(* IEC 61131-3 sources: STAR-PLC-Agent/results/raw/four_group_20261114/star_deepseek_v2/PUB008/functional/attempt_0001, 1 file *)

(* ---- test_program.st ---- *)
PROGRAM PLC_PRG
VAR
 BenchStep : UDINT := 0;
 BenchCalls : UDINT := 0;
 BenchDone : BOOL := FALSE;
 BenchUut0 : FB_Task;
 BenchUut1 : FB_Task;
 BenchUut2 : FB_Task;
 BenchUut3 : FB_Task;
 BenchUut4 : FB_Task;
 BenchUut5 : FB_Task;
 BenchUut6 : FB_Task;
 BenchUut7 : FB_Task;
 BenchUut8 : FB_Task;
 Binding_0_analogValues : ARRAY[-2..4] OF INT;
 Binding_0_channels : ARRAY[7..13] OF ST_AnalogChannel;
 Binding_1_analogValues : ARRAY[1..5] OF INT;
 Binding_1_channels : ARRAY[1..5] OF ST_AnalogChannel;
 Binding_2_analogValues : ARRAY[1..1] OF INT;
 Binding_2_channels : ARRAY[1..1] OF ST_AnalogChannel;
 Binding_3_analogValues : ARRAY[-3..-3] OF INT;
 Binding_3_channels : ARRAY[9..10] OF ST_AnalogChannel;
 Binding_4_analogValues : ARRAY[-3..-1] OF INT;
 Binding_4_channels : ARRAY[7..9] OF ST_AnalogChannel;
 Binding_5_analogValues : ARRAY[-3..0] OF INT;
 Binding_5_channels : ARRAY[8..9] OF ST_AnalogChannel;
 Binding_6_analogValues : ARRAY[-3..-2] OF INT;
 Binding_6_channels : ARRAY[8..11] OF ST_AnalogChannel;
 Binding_7_analogValues : ARRAY[1..5] OF INT;
 Binding_7_channels : ARRAY[1..5] OF ST_AnalogChannel;
 Binding_8_analogValues : ARRAY[1..5] OF INT;
 Binding_8_channels : ARRAY[1..6] OF ST_AnalogChannel;
 TraceIn_count : ARRAY[0..11] OF DINT;
 TraceOut_analogValues_1 : ARRAY[0..11] OF INT;
 TraceOut_analogValues_2 : ARRAY[0..11] OF INT;
 TraceOut_analogValues_3 : ARRAY[0..11] OF INT;
 TraceOut_analogValues_4 : ARRAY[0..11] OF INT;
 TraceOut_analogValues_5 : ARRAY[0..11] OF INT;
 TraceOut_analogValues_6 : ARRAY[0..11] OF INT;
 TraceOut_analogValues_7 : ARRAY[0..11] OF INT;
 TraceOut_channels_1_enable : ARRAY[0..11] OF BOOL;
 TraceOut_channels_1_hiLIM : ARRAY[0..11] OF REAL;
 TraceOut_channels_1_loLIM : ARRAY[0..11] OF REAL;
 TraceOut_channels_1_bipolar : ARRAY[0..11] OF BOOL;
 TraceOut_channels_1_measuringMode : ARRAY[0..11] OF INT;
 TraceOut_channels_1_retVal : ARRAY[0..11] OF WORD;
 TraceOut_channels_1_outputValue : ARRAY[0..11] OF REAL;
 TraceOut_channels_2_enable : ARRAY[0..11] OF BOOL;
 TraceOut_channels_2_hiLIM : ARRAY[0..11] OF REAL;
 TraceOut_channels_2_loLIM : ARRAY[0..11] OF REAL;
 TraceOut_channels_2_bipolar : ARRAY[0..11] OF BOOL;
 TraceOut_channels_2_measuringMode : ARRAY[0..11] OF INT;
 TraceOut_channels_2_retVal : ARRAY[0..11] OF WORD;
 TraceOut_channels_2_outputValue : ARRAY[0..11] OF REAL;
 TraceOut_channels_3_enable : ARRAY[0..11] OF BOOL;
 TraceOut_channels_3_hiLIM : ARRAY[0..11] OF REAL;
 TraceOut_channels_3_loLIM : ARRAY[0..11] OF REAL;
 TraceOut_channels_3_bipolar : ARRAY[0..11] OF BOOL;
 TraceOut_channels_3_measuringMode : ARRAY[0..11] OF INT;
 TraceOut_channels_3_retVal : ARRAY[0..11] OF WORD;
 TraceOut_channels_3_outputValue : ARRAY[0..11] OF REAL;
 TraceOut_channels_4_enable : ARRAY[0..11] OF BOOL;
 TraceOut_channels_4_hiLIM : ARRAY[0..11] OF REAL;
 TraceOut_channels_4_loLIM : ARRAY[0..11] OF REAL;
 TraceOut_channels_4_bipolar : ARRAY[0..11] OF BOOL;
 TraceOut_channels_4_measuringMode : ARRAY[0..11] OF INT;
 TraceOut_channels_4_retVal : ARRAY[0..11] OF WORD;
 TraceOut_channels_4_outputValue : ARRAY[0..11] OF REAL;
 TraceOut_channels_5_enable : ARRAY[0..11] OF BOOL;
 TraceOut_channels_5_hiLIM : ARRAY[0..11] OF REAL;
 TraceOut_channels_5_loLIM : ARRAY[0..11] OF REAL;
 TraceOut_channels_5_bipolar : ARRAY[0..11] OF BOOL;
 TraceOut_channels_5_measuringMode : ARRAY[0..11] OF INT;
 TraceOut_channels_5_retVal : ARRAY[0..11] OF WORD;
 TraceOut_channels_5_outputValue : ARRAY[0..11] OF REAL;
 TraceOut_channels_6_enable : ARRAY[0..11] OF BOOL;
 TraceOut_channels_6_hiLIM : ARRAY[0..11] OF REAL;
 TraceOut_channels_6_loLIM : ARRAY[0..11] OF REAL;
 TraceOut_channels_6_bipolar : ARRAY[0..11] OF BOOL;
 TraceOut_channels_6_measuringMode : ARRAY[0..11] OF INT;
 TraceOut_channels_6_retVal : ARRAY[0..11] OF WORD;
 TraceOut_channels_6_outputValue : ARRAY[0..11] OF REAL;
 TraceOut_channels_7_enable : ARRAY[0..11] OF BOOL;
 TraceOut_channels_7_hiLIM : ARRAY[0..11] OF REAL;
 TraceOut_channels_7_loLIM : ARRAY[0..11] OF REAL;
 TraceOut_channels_7_bipolar : ARRAY[0..11] OF BOOL;
 TraceOut_channels_7_measuringMode : ARRAY[0..11] OF INT;
 TraceOut_channels_7_retVal : ARRAY[0..11] OF WORD;
 TraceOut_channels_7_outputValue : ARRAY[0..11] OF REAL;
END_VAR

IF NOT BenchDone THEN
 CASE BenchStep OF
 0:
   Binding_0_analogValues[-2] := INT#0;
   Binding_0_analogValues[-1] := INT#27648;
   Binding_0_analogValues[0] := INT#-27648;
   Binding_0_analogValues[1] := INT#0;
   Binding_0_analogValues[2] := INT#27648;
   Binding_0_analogValues[3] := INT#1234;
   Binding_0_analogValues[4] := INT#-1234;
   Binding_0_channels[7].enable := TRUE;
   Binding_0_channels[7].hiLIM := REAL#100.0;
   Binding_0_channels[7].loLIM := REAL#0.0;
   Binding_0_channels[7].bipolar := FALSE;
   Binding_0_channels[7].measuringMode := INT#0;
   Binding_0_channels[7].retVal := WORD#7;
   Binding_0_channels[7].outputValue := REAL#-999.0;
   Binding_0_channels[8].enable := TRUE;
   Binding_0_channels[8].hiLIM := REAL#100.0;
   Binding_0_channels[8].loLIM := REAL#0.0;
   Binding_0_channels[8].bipolar := FALSE;
   Binding_0_channels[8].measuringMode := INT#0;
   Binding_0_channels[8].retVal := WORD#7;
   Binding_0_channels[8].outputValue := REAL#-999.0;
   Binding_0_channels[9].enable := TRUE;
   Binding_0_channels[9].hiLIM := REAL#100.0;
   Binding_0_channels[9].loLIM := REAL#0.0;
   Binding_0_channels[9].bipolar := TRUE;
   Binding_0_channels[9].measuringMode := INT#0;
   Binding_0_channels[9].retVal := WORD#7;
   Binding_0_channels[9].outputValue := REAL#-999.0;
   Binding_0_channels[10].enable := TRUE;
   Binding_0_channels[10].hiLIM := REAL#100.0;
   Binding_0_channels[10].loLIM := REAL#0.0;
   Binding_0_channels[10].bipolar := TRUE;
   Binding_0_channels[10].measuringMode := INT#0;
   Binding_0_channels[10].retVal := WORD#7;
   Binding_0_channels[10].outputValue := REAL#-999.0;
   Binding_0_channels[11].enable := TRUE;
   Binding_0_channels[11].hiLIM := REAL#100.0;
   Binding_0_channels[11].loLIM := REAL#0.0;
   Binding_0_channels[11].bipolar := TRUE;
   Binding_0_channels[11].measuringMode := INT#0;
   Binding_0_channels[11].retVal := WORD#7;
   Binding_0_channels[11].outputValue := REAL#-999.0;
   Binding_0_channels[12].enable := TRUE;
   Binding_0_channels[12].hiLIM := REAL#100.0;
   Binding_0_channels[12].loLIM := REAL#0.0;
   Binding_0_channels[12].bipolar := FALSE;
   Binding_0_channels[12].measuringMode := INT#1;
   Binding_0_channels[12].retVal := WORD#7;
   Binding_0_channels[12].outputValue := REAL#-999.0;
   Binding_0_channels[13].enable := TRUE;
   Binding_0_channels[13].hiLIM := REAL#100.0;
   Binding_0_channels[13].loLIM := REAL#0.0;
   Binding_0_channels[13].bipolar := FALSE;
   Binding_0_channels[13].measuringMode := INT#2;
   Binding_0_channels[13].retVal := WORD#7;
   Binding_0_channels[13].outputValue := REAL#-999.0;
   BenchUut0.count := DINT#7;
   TraceIn_count[0] := BenchUut0.count;
   BenchUut0(analogValues := Binding_0_analogValues, channels := Binding_0_channels);
   TraceOut_analogValues_1[0] := Binding_0_analogValues[-2];
   TraceOut_analogValues_2[0] := Binding_0_analogValues[-1];
   TraceOut_analogValues_3[0] := Binding_0_analogValues[0];
   TraceOut_analogValues_4[0] := Binding_0_analogValues[1];
   TraceOut_analogValues_5[0] := Binding_0_analogValues[2];
   TraceOut_analogValues_6[0] := Binding_0_analogValues[3];
   TraceOut_analogValues_7[0] := Binding_0_analogValues[4];
   TraceOut_channels_1_enable[0] := Binding_0_channels[7].enable;
   TraceOut_channels_1_hiLIM[0] := Binding_0_channels[7].hiLIM;
   TraceOut_channels_1_loLIM[0] := Binding_0_channels[7].loLIM;
   TraceOut_channels_1_bipolar[0] := Binding_0_channels[7].bipolar;
   TraceOut_channels_1_measuringMode[0] := Binding_0_channels[7].measuringMode;
   TraceOut_channels_1_retVal[0] := Binding_0_channels[7].retVal;
   TraceOut_channels_1_outputValue[0] := Binding_0_channels[7].outputValue;
   TraceOut_channels_2_enable[0] := Binding_0_channels[8].enable;
   TraceOut_channels_2_hiLIM[0] := Binding_0_channels[8].hiLIM;
   TraceOut_channels_2_loLIM[0] := Binding_0_channels[8].loLIM;
   TraceOut_channels_2_bipolar[0] := Binding_0_channels[8].bipolar;
   TraceOut_channels_2_measuringMode[0] := Binding_0_channels[8].measuringMode;
   TraceOut_channels_2_retVal[0] := Binding_0_channels[8].retVal;
   TraceOut_channels_2_outputValue[0] := Binding_0_channels[8].outputValue;
   TraceOut_channels_3_enable[0] := Binding_0_channels[9].enable;
   TraceOut_channels_3_hiLIM[0] := Binding_0_channels[9].hiLIM;
   TraceOut_channels_3_loLIM[0] := Binding_0_channels[9].loLIM;
   TraceOut_channels_3_bipolar[0] := Binding_0_channels[9].bipolar;
   TraceOut_channels_3_measuringMode[0] := Binding_0_channels[9].measuringMode;
   TraceOut_channels_3_retVal[0] := Binding_0_channels[9].retVal;
   TraceOut_channels_3_outputValue[0] := Binding_0_channels[9].outputValue;
   TraceOut_channels_4_enable[0] := Binding_0_channels[10].enable;
   TraceOut_channels_4_hiLIM[0] := Binding_0_channels[10].hiLIM;
   TraceOut_channels_4_loLIM[0] := Binding_0_channels[10].loLIM;
   TraceOut_channels_4_bipolar[0] := Binding_0_channels[10].bipolar;
   TraceOut_channels_4_measuringMode[0] := Binding_0_channels[10].measuringMode;
   TraceOut_channels_4_retVal[0] := Binding_0_channels[10].retVal;
   TraceOut_channels_4_outputValue[0] := Binding_0_channels[10].outputValue;
   TraceOut_channels_5_enable[0] := Binding_0_channels[11].enable;
   TraceOut_channels_5_hiLIM[0] := Binding_0_channels[11].hiLIM;
   TraceOut_channels_5_loLIM[0] := Binding_0_channels[11].loLIM;
   TraceOut_channels_5_bipolar[0] := Binding_0_channels[11].bipolar;
   TraceOut_channels_5_measuringMode[0] := Binding_0_channels[11].measuringMode;
   TraceOut_channels_5_retVal[0] := Binding_0_channels[11].retVal;
   TraceOut_channels_5_outputValue[0] := Binding_0_channels[11].outputValue;
   TraceOut_channels_6_enable[0] := Binding_0_channels[12].enable;
   TraceOut_channels_6_hiLIM[0] := Binding_0_channels[12].hiLIM;
   TraceOut_channels_6_loLIM[0] := Binding_0_channels[12].loLIM;
   TraceOut_channels_6_bipolar[0] := Binding_0_channels[12].bipolar;
   TraceOut_channels_6_measuringMode[0] := Binding_0_channels[12].measuringMode;
   TraceOut_channels_6_retVal[0] := Binding_0_channels[12].retVal;
   TraceOut_channels_6_outputValue[0] := Binding_0_channels[12].outputValue;
   TraceOut_channels_7_enable[0] := Binding_0_channels[13].enable;
   TraceOut_channels_7_hiLIM[0] := Binding_0_channels[13].hiLIM;
   TraceOut_channels_7_loLIM[0] := Binding_0_channels[13].loLIM;
   TraceOut_channels_7_bipolar[0] := Binding_0_channels[13].bipolar;
   TraceOut_channels_7_measuringMode[0] := Binding_0_channels[13].measuringMode;
   TraceOut_channels_7_retVal[0] := Binding_0_channels[13].retVal;
   TraceOut_channels_7_outputValue[0] := Binding_0_channels[13].outputValue;
   BenchCalls := BenchCalls + 1;
 1:
   Binding_1_analogValues[1] := INT#1;
   Binding_1_analogValues[2] := INT#2;
   Binding_1_analogValues[3] := INT#3;
   Binding_1_analogValues[4] := INT#4;
   Binding_1_analogValues[5] := INT#5;
   Binding_1_channels[1].enable := FALSE;
   Binding_1_channels[1].hiLIM := REAL#100.0;
   Binding_1_channels[1].loLIM := REAL#0.0;
   Binding_1_channels[1].bipolar := FALSE;
   Binding_1_channels[1].measuringMode := INT#0;
   Binding_1_channels[1].retVal := WORD#7;
   Binding_1_channels[1].outputValue := REAL#-999.0;
   Binding_1_channels[2].enable := TRUE;
   Binding_1_channels[2].hiLIM := REAL#0.0;
   Binding_1_channels[2].loLIM := REAL#10.0;
   Binding_1_channels[2].bipolar := FALSE;
   Binding_1_channels[2].measuringMode := INT#9;
   Binding_1_channels[2].retVal := WORD#7;
   Binding_1_channels[2].outputValue := REAL#-999.0;
   Binding_1_channels[3].enable := TRUE;
   Binding_1_channels[3].hiLIM := REAL#10.0;
   Binding_1_channels[3].loLIM := REAL#10.0;
   Binding_1_channels[3].bipolar := FALSE;
   Binding_1_channels[3].measuringMode := INT#0;
   Binding_1_channels[3].retVal := WORD#7;
   Binding_1_channels[3].outputValue := REAL#-999.0;
   Binding_1_channels[4].enable := TRUE;
   Binding_1_channels[4].hiLIM := REAL#100.0;
   Binding_1_channels[4].loLIM := REAL#0.0;
   Binding_1_channels[4].bipolar := FALSE;
   Binding_1_channels[4].measuringMode := INT#2;
   Binding_1_channels[4].retVal := WORD#7;
   Binding_1_channels[4].outputValue := REAL#-999.0;
   Binding_1_channels[5].enable := TRUE;
   Binding_1_channels[5].hiLIM := REAL#100.0;
   Binding_1_channels[5].loLIM := REAL#0.0;
   Binding_1_channels[5].bipolar := FALSE;
   Binding_1_channels[5].measuringMode := INT#0;
   Binding_1_channels[5].retVal := WORD#7;
   Binding_1_channels[5].outputValue := REAL#-999.0;
   BenchUut1.count := DINT#4;
   TraceIn_count[1] := BenchUut1.count;
   BenchUut1(analogValues := Binding_1_analogValues, channels := Binding_1_channels);
   TraceOut_analogValues_1[1] := Binding_1_analogValues[1];
   TraceOut_analogValues_2[1] := Binding_1_analogValues[2];
   TraceOut_analogValues_3[1] := Binding_1_analogValues[3];
   TraceOut_analogValues_4[1] := Binding_1_analogValues[4];
   TraceOut_analogValues_5[1] := Binding_1_analogValues[5];
   TraceOut_channels_1_enable[1] := Binding_1_channels[1].enable;
   TraceOut_channels_1_hiLIM[1] := Binding_1_channels[1].hiLIM;
   TraceOut_channels_1_loLIM[1] := Binding_1_channels[1].loLIM;
   TraceOut_channels_1_bipolar[1] := Binding_1_channels[1].bipolar;
   TraceOut_channels_1_measuringMode[1] := Binding_1_channels[1].measuringMode;
   TraceOut_channels_1_retVal[1] := Binding_1_channels[1].retVal;
   TraceOut_channels_1_outputValue[1] := Binding_1_channels[1].outputValue;
   TraceOut_channels_2_enable[1] := Binding_1_channels[2].enable;
   TraceOut_channels_2_hiLIM[1] := Binding_1_channels[2].hiLIM;
   TraceOut_channels_2_loLIM[1] := Binding_1_channels[2].loLIM;
   TraceOut_channels_2_bipolar[1] := Binding_1_channels[2].bipolar;
   TraceOut_channels_2_measuringMode[1] := Binding_1_channels[2].measuringMode;
   TraceOut_channels_2_retVal[1] := Binding_1_channels[2].retVal;
   TraceOut_channels_2_outputValue[1] := Binding_1_channels[2].outputValue;
   TraceOut_channels_3_enable[1] := Binding_1_channels[3].enable;
   TraceOut_channels_3_hiLIM[1] := Binding_1_channels[3].hiLIM;
   TraceOut_channels_3_loLIM[1] := Binding_1_channels[3].loLIM;
   TraceOut_channels_3_bipolar[1] := Binding_1_channels[3].bipolar;
   TraceOut_channels_3_measuringMode[1] := Binding_1_channels[3].measuringMode;
   TraceOut_channels_3_retVal[1] := Binding_1_channels[3].retVal;
   TraceOut_channels_3_outputValue[1] := Binding_1_channels[3].outputValue;
   TraceOut_channels_4_enable[1] := Binding_1_channels[4].enable;
   TraceOut_channels_4_hiLIM[1] := Binding_1_channels[4].hiLIM;
   TraceOut_channels_4_loLIM[1] := Binding_1_channels[4].loLIM;
   TraceOut_channels_4_bipolar[1] := Binding_1_channels[4].bipolar;
   TraceOut_channels_4_measuringMode[1] := Binding_1_channels[4].measuringMode;
   TraceOut_channels_4_retVal[1] := Binding_1_channels[4].retVal;
   TraceOut_channels_4_outputValue[1] := Binding_1_channels[4].outputValue;
   TraceOut_channels_5_enable[1] := Binding_1_channels[5].enable;
   TraceOut_channels_5_hiLIM[1] := Binding_1_channels[5].hiLIM;
   TraceOut_channels_5_loLIM[1] := Binding_1_channels[5].loLIM;
   TraceOut_channels_5_bipolar[1] := Binding_1_channels[5].bipolar;
   TraceOut_channels_5_measuringMode[1] := Binding_1_channels[5].measuringMode;
   TraceOut_channels_5_retVal[1] := Binding_1_channels[5].retVal;
   TraceOut_channels_5_outputValue[1] := Binding_1_channels[5].outputValue;
   BenchCalls := BenchCalls + 1;
 2:
   Binding_2_analogValues[1] := INT#-27648;
   Binding_2_channels[1].enable := TRUE;
   Binding_2_channels[1].hiLIM := REAL#100.0;
   Binding_2_channels[1].loLIM := REAL#0.0;
   Binding_2_channels[1].bipolar := FALSE;
   Binding_2_channels[1].measuringMode := INT#0;
   Binding_2_channels[1].retVal := WORD#7;
   Binding_2_channels[1].outputValue := REAL#-999.0;
   BenchUut2.count := DINT#0;
   TraceIn_count[2] := BenchUut2.count;
   BenchUut2(analogValues := Binding_2_analogValues, channels := Binding_2_channels);
   TraceOut_analogValues_1[2] := Binding_2_analogValues[1];
   TraceOut_channels_1_enable[2] := Binding_2_channels[1].enable;
   TraceOut_channels_1_hiLIM[2] := Binding_2_channels[1].hiLIM;
   TraceOut_channels_1_loLIM[2] := Binding_2_channels[1].loLIM;
   TraceOut_channels_1_bipolar[2] := Binding_2_channels[1].bipolar;
   TraceOut_channels_1_measuringMode[2] := Binding_2_channels[1].measuringMode;
   TraceOut_channels_1_retVal[2] := Binding_2_channels[1].retVal;
   TraceOut_channels_1_outputValue[2] := Binding_2_channels[1].outputValue;
   BenchCalls := BenchCalls + 1;
 3:
   Binding_2_analogValues[1] := INT#-27648;
   Binding_2_channels[1].enable := TRUE;
   Binding_2_channels[1].hiLIM := REAL#100.0;
   Binding_2_channels[1].loLIM := REAL#0.0;
   Binding_2_channels[1].bipolar := FALSE;
   Binding_2_channels[1].measuringMode := INT#0;
   Binding_2_channels[1].retVal := WORD#7;
   Binding_2_channels[1].outputValue := REAL#-999.0;
   BenchUut2.count := DINT#1;
   TraceIn_count[3] := BenchUut2.count;
   BenchUut2(analogValues := Binding_2_analogValues, channels := Binding_2_channels);
   TraceOut_analogValues_1[3] := Binding_2_analogValues[1];
   TraceOut_channels_1_enable[3] := Binding_2_channels[1].enable;
   TraceOut_channels_1_hiLIM[3] := Binding_2_channels[1].hiLIM;
   TraceOut_channels_1_loLIM[3] := Binding_2_channels[1].loLIM;
   TraceOut_channels_1_bipolar[3] := Binding_2_channels[1].bipolar;
   TraceOut_channels_1_measuringMode[3] := Binding_2_channels[1].measuringMode;
   TraceOut_channels_1_retVal[3] := Binding_2_channels[1].retVal;
   TraceOut_channels_1_outputValue[3] := Binding_2_channels[1].outputValue;
   BenchCalls := BenchCalls + 1;
 4:
   Binding_3_analogValues[-3] := INT#32767;
   Binding_3_channels[9].enable := TRUE;
   Binding_3_channels[9].hiLIM := REAL#27648.0;
   Binding_3_channels[9].loLIM := REAL#-27648.0;
   Binding_3_channels[9].bipolar := TRUE;
   Binding_3_channels[9].measuringMode := INT#0;
   Binding_3_channels[9].retVal := WORD#7;
   Binding_3_channels[9].outputValue := REAL#-999.0;
   Binding_3_channels[10].enable := TRUE;
   Binding_3_channels[10].hiLIM := REAL#27648.0;
   Binding_3_channels[10].loLIM := REAL#-27648.0;
   Binding_3_channels[10].bipolar := TRUE;
   Binding_3_channels[10].measuringMode := INT#0;
   Binding_3_channels[10].retVal := WORD#7;
   Binding_3_channels[10].outputValue := REAL#33.0;
   BenchUut3.count := DINT#1;
   TraceIn_count[4] := BenchUut3.count;
   BenchUut3(analogValues := Binding_3_analogValues, channels := Binding_3_channels);
   TraceOut_analogValues_1[4] := Binding_3_analogValues[-3];
   TraceOut_channels_1_enable[4] := Binding_3_channels[9].enable;
   TraceOut_channels_1_hiLIM[4] := Binding_3_channels[9].hiLIM;
   TraceOut_channels_1_loLIM[4] := Binding_3_channels[9].loLIM;
   TraceOut_channels_1_bipolar[4] := Binding_3_channels[9].bipolar;
   TraceOut_channels_1_measuringMode[4] := Binding_3_channels[9].measuringMode;
   TraceOut_channels_1_retVal[4] := Binding_3_channels[9].retVal;
   TraceOut_channels_1_outputValue[4] := Binding_3_channels[9].outputValue;
   TraceOut_channels_2_enable[4] := Binding_3_channels[10].enable;
   TraceOut_channels_2_hiLIM[4] := Binding_3_channels[10].hiLIM;
   TraceOut_channels_2_loLIM[4] := Binding_3_channels[10].loLIM;
   TraceOut_channels_2_bipolar[4] := Binding_3_channels[10].bipolar;
   TraceOut_channels_2_measuringMode[4] := Binding_3_channels[10].measuringMode;
   TraceOut_channels_2_retVal[4] := Binding_3_channels[10].retVal;
   TraceOut_channels_2_outputValue[4] := Binding_3_channels[10].outputValue;
   BenchCalls := BenchCalls + 1;
 5:
   Binding_4_analogValues[-3] := INT#1000;
   Binding_4_analogValues[-2] := INT#-1000;
   Binding_4_analogValues[-1] := INT#30000;
   Binding_4_channels[7].enable := FALSE;
   Binding_4_channels[7].hiLIM := REAL#0.0;
   Binding_4_channels[7].loLIM := REAL#100.0;
   Binding_4_channels[7].bipolar := FALSE;
   Binding_4_channels[7].measuringMode := INT#9;
   Binding_4_channels[7].retVal := WORD#123;
   Binding_4_channels[7].outputValue := REAL#-42.5;
   Binding_4_channels[8].enable := TRUE;
   Binding_4_channels[8].hiLIM := REAL#5.0;
   Binding_4_channels[8].loLIM := REAL#5.0;
   Binding_4_channels[8].bipolar := FALSE;
   Binding_4_channels[8].measuringMode := INT#1;
   Binding_4_channels[8].retVal := WORD#0;
   Binding_4_channels[8].outputValue := REAL#12.25;
   Binding_4_channels[9].enable := TRUE;
   Binding_4_channels[9].hiLIM := REAL#100.0;
   Binding_4_channels[9].loLIM := REAL#0.0;
   Binding_4_channels[9].bipolar := FALSE;
   Binding_4_channels[9].measuringMode := INT#0;
   Binding_4_channels[9].retVal := WORD#0;
   Binding_4_channels[9].outputValue := REAL#0.0;
   BenchUut4.count := DINT#3;
   TraceIn_count[5] := BenchUut4.count;
   BenchUut4(analogValues := Binding_4_analogValues, channels := Binding_4_channels);
   TraceOut_analogValues_1[5] := Binding_4_analogValues[-3];
   TraceOut_analogValues_2[5] := Binding_4_analogValues[-2];
   TraceOut_analogValues_3[5] := Binding_4_analogValues[-1];
   TraceOut_channels_1_enable[5] := Binding_4_channels[7].enable;
   TraceOut_channels_1_hiLIM[5] := Binding_4_channels[7].hiLIM;
   TraceOut_channels_1_loLIM[5] := Binding_4_channels[7].loLIM;
   TraceOut_channels_1_bipolar[5] := Binding_4_channels[7].bipolar;
   TraceOut_channels_1_measuringMode[5] := Binding_4_channels[7].measuringMode;
   TraceOut_channels_1_retVal[5] := Binding_4_channels[7].retVal;
   TraceOut_channels_1_outputValue[5] := Binding_4_channels[7].outputValue;
   TraceOut_channels_2_enable[5] := Binding_4_channels[8].enable;
   TraceOut_channels_2_hiLIM[5] := Binding_4_channels[8].hiLIM;
   TraceOut_channels_2_loLIM[5] := Binding_4_channels[8].loLIM;
   TraceOut_channels_2_bipolar[5] := Binding_4_channels[8].bipolar;
   TraceOut_channels_2_measuringMode[5] := Binding_4_channels[8].measuringMode;
   TraceOut_channels_2_retVal[5] := Binding_4_channels[8].retVal;
   TraceOut_channels_2_outputValue[5] := Binding_4_channels[8].outputValue;
   TraceOut_channels_3_enable[5] := Binding_4_channels[9].enable;
   TraceOut_channels_3_hiLIM[5] := Binding_4_channels[9].hiLIM;
   TraceOut_channels_3_loLIM[5] := Binding_4_channels[9].loLIM;
   TraceOut_channels_3_bipolar[5] := Binding_4_channels[9].bipolar;
   TraceOut_channels_3_measuringMode[5] := Binding_4_channels[9].measuringMode;
   TraceOut_channels_3_retVal[5] := Binding_4_channels[9].retVal;
   TraceOut_channels_3_outputValue[5] := Binding_4_channels[9].outputValue;
   BenchCalls := BenchCalls + 1;
 6:
   Binding_4_analogValues[-3] := INT#-30000;
   Binding_4_analogValues[-2] := INT#1234;
   Binding_4_analogValues[-1] := INT#0;
   Binding_4_analogValues[0] := INT#999;
   Binding_4_channels[7].enable := TRUE;
   Binding_4_channels[7].hiLIM := REAL#10.0;
   Binding_4_channels[7].loLIM := REAL#-10.0;
   Binding_4_channels[7].bipolar := FALSE;
   Binding_4_channels[7].measuringMode := INT#2;
   Binding_4_channels[7].retVal := WORD#0;
   Binding_4_channels[7].outputValue := REAL#1.0;
   Binding_4_channels[8].enable := TRUE;
   Binding_4_channels[8].hiLIM := REAL#10.0;
   Binding_4_channels[8].loLIM := REAL#20.0;
   Binding_4_channels[8].bipolar := FALSE;
   Binding_4_channels[8].measuringMode := INT#2;
   Binding_4_channels[8].retVal := WORD#0;
   Binding_4_channels[8].outputValue := REAL#3.5;
   Binding_4_channels[9].enable := TRUE;
   Binding_4_channels[9].hiLIM := REAL#10.0;
   Binding_4_channels[9].loLIM := REAL#0.0;
   Binding_4_channels[9].bipolar := TRUE;
   Binding_4_channels[9].measuringMode := INT#0;
   Binding_4_channels[9].retVal := WORD#0;
   Binding_4_channels[9].outputValue := REAL#0.0;
   BenchUut4.count := DINT#3;
   TraceIn_count[6] := BenchUut4.count;
   BenchUut4(analogValues := Binding_4_analogValues, channels := Binding_4_channels);
   TraceOut_analogValues_1[6] := Binding_4_analogValues[-3];
   TraceOut_analogValues_2[6] := Binding_4_analogValues[-2];
   TraceOut_analogValues_3[6] := Binding_4_analogValues[-1];
   TraceOut_analogValues_4[6] := Binding_4_analogValues[0];
   TraceOut_channels_1_enable[6] := Binding_4_channels[7].enable;
   TraceOut_channels_1_hiLIM[6] := Binding_4_channels[7].hiLIM;
   TraceOut_channels_1_loLIM[6] := Binding_4_channels[7].loLIM;
   TraceOut_channels_1_bipolar[6] := Binding_4_channels[7].bipolar;
   TraceOut_channels_1_measuringMode[6] := Binding_4_channels[7].measuringMode;
   TraceOut_channels_1_retVal[6] := Binding_4_channels[7].retVal;
   TraceOut_channels_1_outputValue[6] := Binding_4_channels[7].outputValue;
   TraceOut_channels_2_enable[6] := Binding_4_channels[8].enable;
   TraceOut_channels_2_hiLIM[6] := Binding_4_channels[8].hiLIM;
   TraceOut_channels_2_loLIM[6] := Binding_4_channels[8].loLIM;
   TraceOut_channels_2_bipolar[6] := Binding_4_channels[8].bipolar;
   TraceOut_channels_2_measuringMode[6] := Binding_4_channels[8].measuringMode;
   TraceOut_channels_2_retVal[6] := Binding_4_channels[8].retVal;
   TraceOut_channels_2_outputValue[6] := Binding_4_channels[8].outputValue;
   TraceOut_channels_3_enable[6] := Binding_4_channels[9].enable;
   TraceOut_channels_3_hiLIM[6] := Binding_4_channels[9].hiLIM;
   TraceOut_channels_3_loLIM[6] := Binding_4_channels[9].loLIM;
   TraceOut_channels_3_bipolar[6] := Binding_4_channels[9].bipolar;
   TraceOut_channels_3_measuringMode[6] := Binding_4_channels[9].measuringMode;
   TraceOut_channels_3_retVal[6] := Binding_4_channels[9].retVal;
   TraceOut_channels_3_outputValue[6] := Binding_4_channels[9].outputValue;
   BenchCalls := BenchCalls + 1;
 7:
   Binding_5_analogValues[-3] := INT#0;
   Binding_5_analogValues[-2] := INT#27648;
   Binding_5_analogValues[-1] := INT#-27648;
   Binding_5_analogValues[0] := INT#0;
   Binding_5_channels[8].enable := TRUE;
   Binding_5_channels[8].hiLIM := REAL#100.0;
   Binding_5_channels[8].loLIM := REAL#0.0;
   Binding_5_channels[8].bipolar := FALSE;
   Binding_5_channels[8].measuringMode := INT#0;
   Binding_5_channels[8].retVal := WORD#7;
   Binding_5_channels[8].outputValue := REAL#-999.0;
   Binding_5_channels[9].enable := TRUE;
   Binding_5_channels[9].hiLIM := REAL#100.0;
   Binding_5_channels[9].loLIM := REAL#0.0;
   Binding_5_channels[9].bipolar := FALSE;
   Binding_5_channels[9].measuringMode := INT#0;
   Binding_5_channels[9].retVal := WORD#7;
   Binding_5_channels[9].outputValue := REAL#-999.0;
   BenchUut5.count := DINT#2;
   TraceIn_count[7] := BenchUut5.count;
   BenchUut5(analogValues := Binding_5_analogValues, channels := Binding_5_channels);
   TraceOut_analogValues_1[7] := Binding_5_analogValues[-3];
   TraceOut_analogValues_2[7] := Binding_5_analogValues[-2];
   TraceOut_analogValues_3[7] := Binding_5_analogValues[-1];
   TraceOut_analogValues_4[7] := Binding_5_analogValues[0];
   TraceOut_channels_1_enable[7] := Binding_5_channels[8].enable;
   TraceOut_channels_1_hiLIM[7] := Binding_5_channels[8].hiLIM;
   TraceOut_channels_1_loLIM[7] := Binding_5_channels[8].loLIM;
   TraceOut_channels_1_bipolar[7] := Binding_5_channels[8].bipolar;
   TraceOut_channels_1_measuringMode[7] := Binding_5_channels[8].measuringMode;
   TraceOut_channels_1_retVal[7] := Binding_5_channels[8].retVal;
   TraceOut_channels_1_outputValue[7] := Binding_5_channels[8].outputValue;
   TraceOut_channels_2_enable[7] := Binding_5_channels[9].enable;
   TraceOut_channels_2_hiLIM[7] := Binding_5_channels[9].hiLIM;
   TraceOut_channels_2_loLIM[7] := Binding_5_channels[9].loLIM;
   TraceOut_channels_2_bipolar[7] := Binding_5_channels[9].bipolar;
   TraceOut_channels_2_measuringMode[7] := Binding_5_channels[9].measuringMode;
   TraceOut_channels_2_retVal[7] := Binding_5_channels[9].retVal;
   TraceOut_channels_2_outputValue[7] := Binding_5_channels[9].outputValue;
   BenchCalls := BenchCalls + 1;
 8:
   Binding_6_analogValues[-3] := INT#0;
   Binding_6_analogValues[-2] := INT#27648;
   Binding_6_channels[8].enable := TRUE;
   Binding_6_channels[8].hiLIM := REAL#100.0;
   Binding_6_channels[8].loLIM := REAL#0.0;
   Binding_6_channels[8].bipolar := FALSE;
   Binding_6_channels[8].measuringMode := INT#0;
   Binding_6_channels[8].retVal := WORD#7;
   Binding_6_channels[8].outputValue := REAL#-999.0;
   Binding_6_channels[9].enable := TRUE;
   Binding_6_channels[9].hiLIM := REAL#100.0;
   Binding_6_channels[9].loLIM := REAL#0.0;
   Binding_6_channels[9].bipolar := FALSE;
   Binding_6_channels[9].measuringMode := INT#0;
   Binding_6_channels[9].retVal := WORD#7;
   Binding_6_channels[9].outputValue := REAL#-999.0;
   Binding_6_channels[10].enable := TRUE;
   Binding_6_channels[10].hiLIM := REAL#100.0;
   Binding_6_channels[10].loLIM := REAL#0.0;
   Binding_6_channels[10].bipolar := TRUE;
   Binding_6_channels[10].measuringMode := INT#0;
   Binding_6_channels[10].retVal := WORD#7;
   Binding_6_channels[10].outputValue := REAL#-999.0;
   Binding_6_channels[11].enable := TRUE;
   Binding_6_channels[11].hiLIM := REAL#100.0;
   Binding_6_channels[11].loLIM := REAL#0.0;
   Binding_6_channels[11].bipolar := TRUE;
   Binding_6_channels[11].measuringMode := INT#0;
   Binding_6_channels[11].retVal := WORD#7;
   Binding_6_channels[11].outputValue := REAL#-999.0;
   BenchUut6.count := DINT#2;
   TraceIn_count[8] := BenchUut6.count;
   BenchUut6(analogValues := Binding_6_analogValues, channels := Binding_6_channels);
   TraceOut_analogValues_1[8] := Binding_6_analogValues[-3];
   TraceOut_analogValues_2[8] := Binding_6_analogValues[-2];
   TraceOut_channels_1_enable[8] := Binding_6_channels[8].enable;
   TraceOut_channels_1_hiLIM[8] := Binding_6_channels[8].hiLIM;
   TraceOut_channels_1_loLIM[8] := Binding_6_channels[8].loLIM;
   TraceOut_channels_1_bipolar[8] := Binding_6_channels[8].bipolar;
   TraceOut_channels_1_measuringMode[8] := Binding_6_channels[8].measuringMode;
   TraceOut_channels_1_retVal[8] := Binding_6_channels[8].retVal;
   TraceOut_channels_1_outputValue[8] := Binding_6_channels[8].outputValue;
   TraceOut_channels_2_enable[8] := Binding_6_channels[9].enable;
   TraceOut_channels_2_hiLIM[8] := Binding_6_channels[9].hiLIM;
   TraceOut_channels_2_loLIM[8] := Binding_6_channels[9].loLIM;
   TraceOut_channels_2_bipolar[8] := Binding_6_channels[9].bipolar;
   TraceOut_channels_2_measuringMode[8] := Binding_6_channels[9].measuringMode;
   TraceOut_channels_2_retVal[8] := Binding_6_channels[9].retVal;
   TraceOut_channels_2_outputValue[8] := Binding_6_channels[9].outputValue;
   TraceOut_channels_3_enable[8] := Binding_6_channels[10].enable;
   TraceOut_channels_3_hiLIM[8] := Binding_6_channels[10].hiLIM;
   TraceOut_channels_3_loLIM[8] := Binding_6_channels[10].loLIM;
   TraceOut_channels_3_bipolar[8] := Binding_6_channels[10].bipolar;
   TraceOut_channels_3_measuringMode[8] := Binding_6_channels[10].measuringMode;
   TraceOut_channels_3_retVal[8] := Binding_6_channels[10].retVal;
   TraceOut_channels_3_outputValue[8] := Binding_6_channels[10].outputValue;
   TraceOut_channels_4_enable[8] := Binding_6_channels[11].enable;
   TraceOut_channels_4_hiLIM[8] := Binding_6_channels[11].hiLIM;
   TraceOut_channels_4_loLIM[8] := Binding_6_channels[11].loLIM;
   TraceOut_channels_4_bipolar[8] := Binding_6_channels[11].bipolar;
   TraceOut_channels_4_measuringMode[8] := Binding_6_channels[11].measuringMode;
   TraceOut_channels_4_retVal[8] := Binding_6_channels[11].retVal;
   TraceOut_channels_4_outputValue[8] := Binding_6_channels[11].outputValue;
   BenchCalls := BenchCalls + 1;
 9:
   Binding_7_analogValues[1] := INT#27648;
   Binding_7_analogValues[2] := INT#13824;
   Binding_7_analogValues[3] := INT#27648;
   Binding_7_analogValues[4] := INT#27648;
   Binding_7_analogValues[5] := INT#500;
   Binding_7_channels[1].enable := TRUE;
   Binding_7_channels[1].hiLIM := REAL#100.0;
   Binding_7_channels[1].loLIM := REAL#0.0;
   Binding_7_channels[1].bipolar := FALSE;
   Binding_7_channels[1].measuringMode := INT#0;
   Binding_7_channels[1].retVal := WORD#7;
   Binding_7_channels[1].outputValue := REAL#-999.0;
   Binding_7_channels[2].enable := TRUE;
   Binding_7_channels[2].hiLIM := REAL#50.0;
   Binding_7_channels[2].loLIM := REAL#-50.0;
   Binding_7_channels[2].bipolar := FALSE;
   Binding_7_channels[2].measuringMode := INT#0;
   Binding_7_channels[2].retVal := WORD#7;
   Binding_7_channels[2].outputValue := REAL#-999.0;
   Binding_7_channels[3].enable := TRUE;
   Binding_7_channels[3].hiLIM := REAL#100.0;
   Binding_7_channels[3].loLIM := REAL#0.0;
   Binding_7_channels[3].bipolar := FALSE;
   Binding_7_channels[3].measuringMode := INT#0;
   Binding_7_channels[3].retVal := WORD#7;
   Binding_7_channels[3].outputValue := REAL#-999.0;
   Binding_7_channels[4].enable := TRUE;
   Binding_7_channels[4].hiLIM := REAL#100.0;
   Binding_7_channels[4].loLIM := REAL#0.0;
   Binding_7_channels[4].bipolar := FALSE;
   Binding_7_channels[4].measuringMode := INT#0;
   Binding_7_channels[4].retVal := WORD#7;
   Binding_7_channels[4].outputValue := REAL#-999.0;
   Binding_7_channels[5].enable := TRUE;
   Binding_7_channels[5].hiLIM := REAL#100.0;
   Binding_7_channels[5].loLIM := REAL#0.0;
   Binding_7_channels[5].bipolar := FALSE;
   Binding_7_channels[5].measuringMode := INT#1;
   Binding_7_channels[5].retVal := WORD#7;
   Binding_7_channels[5].outputValue := REAL#-999.0;
   BenchUut7.count := DINT#5;
   TraceIn_count[9] := BenchUut7.count;
   BenchUut7(analogValues := Binding_7_analogValues, channels := Binding_7_channels);
   TraceOut_analogValues_1[9] := Binding_7_analogValues[1];
   TraceOut_analogValues_2[9] := Binding_7_analogValues[2];
   TraceOut_analogValues_3[9] := Binding_7_analogValues[3];
   TraceOut_analogValues_4[9] := Binding_7_analogValues[4];
   TraceOut_analogValues_5[9] := Binding_7_analogValues[5];
   TraceOut_channels_1_enable[9] := Binding_7_channels[1].enable;
   TraceOut_channels_1_hiLIM[9] := Binding_7_channels[1].hiLIM;
   TraceOut_channels_1_loLIM[9] := Binding_7_channels[1].loLIM;
   TraceOut_channels_1_bipolar[9] := Binding_7_channels[1].bipolar;
   TraceOut_channels_1_measuringMode[9] := Binding_7_channels[1].measuringMode;
   TraceOut_channels_1_retVal[9] := Binding_7_channels[1].retVal;
   TraceOut_channels_1_outputValue[9] := Binding_7_channels[1].outputValue;
   TraceOut_channels_2_enable[9] := Binding_7_channels[2].enable;
   TraceOut_channels_2_hiLIM[9] := Binding_7_channels[2].hiLIM;
   TraceOut_channels_2_loLIM[9] := Binding_7_channels[2].loLIM;
   TraceOut_channels_2_bipolar[9] := Binding_7_channels[2].bipolar;
   TraceOut_channels_2_measuringMode[9] := Binding_7_channels[2].measuringMode;
   TraceOut_channels_2_retVal[9] := Binding_7_channels[2].retVal;
   TraceOut_channels_2_outputValue[9] := Binding_7_channels[2].outputValue;
   TraceOut_channels_3_enable[9] := Binding_7_channels[3].enable;
   TraceOut_channels_3_hiLIM[9] := Binding_7_channels[3].hiLIM;
   TraceOut_channels_3_loLIM[9] := Binding_7_channels[3].loLIM;
   TraceOut_channels_3_bipolar[9] := Binding_7_channels[3].bipolar;
   TraceOut_channels_3_measuringMode[9] := Binding_7_channels[3].measuringMode;
   TraceOut_channels_3_retVal[9] := Binding_7_channels[3].retVal;
   TraceOut_channels_3_outputValue[9] := Binding_7_channels[3].outputValue;
   TraceOut_channels_4_enable[9] := Binding_7_channels[4].enable;
   TraceOut_channels_4_hiLIM[9] := Binding_7_channels[4].hiLIM;
   TraceOut_channels_4_loLIM[9] := Binding_7_channels[4].loLIM;
   TraceOut_channels_4_bipolar[9] := Binding_7_channels[4].bipolar;
   TraceOut_channels_4_measuringMode[9] := Binding_7_channels[4].measuringMode;
   TraceOut_channels_4_retVal[9] := Binding_7_channels[4].retVal;
   TraceOut_channels_4_outputValue[9] := Binding_7_channels[4].outputValue;
   TraceOut_channels_5_enable[9] := Binding_7_channels[5].enable;
   TraceOut_channels_5_hiLIM[9] := Binding_7_channels[5].hiLIM;
   TraceOut_channels_5_loLIM[9] := Binding_7_channels[5].loLIM;
   TraceOut_channels_5_bipolar[9] := Binding_7_channels[5].bipolar;
   TraceOut_channels_5_measuringMode[9] := Binding_7_channels[5].measuringMode;
   TraceOut_channels_5_retVal[9] := Binding_7_channels[5].retVal;
   TraceOut_channels_5_outputValue[9] := Binding_7_channels[5].outputValue;
   BenchCalls := BenchCalls + 1;
 10:
   Binding_7_analogValues[1] := INT#0;
   Binding_7_analogValues[2] := INT#0;
   Binding_7_analogValues[3] := INT#0;
   Binding_7_analogValues[4] := INT#0;
   Binding_7_analogValues[5] := INT#9999;
   Binding_7_channels[1].enable := FALSE;
   Binding_7_channels[1].hiLIM := REAL#10.0;
   Binding_7_channels[1].loLIM := REAL#20.0;
   Binding_7_channels[1].bipolar := FALSE;
   Binding_7_channels[1].measuringMode := INT#9;
   Binding_7_channels[1].retVal := WORD#0;
   Binding_7_channels[1].outputValue := REAL#100.0;
   Binding_7_channels[2].enable := TRUE;
   Binding_7_channels[2].hiLIM := REAL#10.0;
   Binding_7_channels[2].loLIM := REAL#20.0;
   Binding_7_channels[2].bipolar := FALSE;
   Binding_7_channels[2].measuringMode := INT#9;
   Binding_7_channels[2].retVal := WORD#0;
   Binding_7_channels[2].outputValue := REAL#0.0;
   Binding_7_channels[3].enable := TRUE;
   Binding_7_channels[3].hiLIM := REAL#10.0;
   Binding_7_channels[3].loLIM := REAL#10.0;
   Binding_7_channels[3].bipolar := FALSE;
   Binding_7_channels[3].measuringMode := INT#0;
   Binding_7_channels[3].retVal := WORD#0;
   Binding_7_channels[3].outputValue := REAL#100.0;
   Binding_7_channels[4].enable := TRUE;
   Binding_7_channels[4].hiLIM := REAL#200.0;
   Binding_7_channels[4].loLIM := REAL#100.0;
   Binding_7_channels[4].bipolar := FALSE;
   Binding_7_channels[4].measuringMode := INT#0;
   Binding_7_channels[4].retVal := WORD#0;
   Binding_7_channels[4].outputValue := REAL#100.0;
   Binding_7_channels[5].enable := TRUE;
   Binding_7_channels[5].hiLIM := REAL#100.0;
   Binding_7_channels[5].loLIM := REAL#0.0;
   Binding_7_channels[5].bipolar := FALSE;
   Binding_7_channels[5].measuringMode := INT#1;
   Binding_7_channels[5].retVal := WORD#0;
   Binding_7_channels[5].outputValue := REAL#50.0;
   BenchUut7.count := DINT#4;
   TraceIn_count[10] := BenchUut7.count;
   BenchUut7(analogValues := Binding_7_analogValues, channels := Binding_7_channels);
   TraceOut_analogValues_1[10] := Binding_7_analogValues[1];
   TraceOut_analogValues_2[10] := Binding_7_analogValues[2];
   TraceOut_analogValues_3[10] := Binding_7_analogValues[3];
   TraceOut_analogValues_4[10] := Binding_7_analogValues[4];
   TraceOut_analogValues_5[10] := Binding_7_analogValues[5];
   TraceOut_channels_1_enable[10] := Binding_7_channels[1].enable;
   TraceOut_channels_1_hiLIM[10] := Binding_7_channels[1].hiLIM;
   TraceOut_channels_1_loLIM[10] := Binding_7_channels[1].loLIM;
   TraceOut_channels_1_bipolar[10] := Binding_7_channels[1].bipolar;
   TraceOut_channels_1_measuringMode[10] := Binding_7_channels[1].measuringMode;
   TraceOut_channels_1_retVal[10] := Binding_7_channels[1].retVal;
   TraceOut_channels_1_outputValue[10] := Binding_7_channels[1].outputValue;
   TraceOut_channels_2_enable[10] := Binding_7_channels[2].enable;
   TraceOut_channels_2_hiLIM[10] := Binding_7_channels[2].hiLIM;
   TraceOut_channels_2_loLIM[10] := Binding_7_channels[2].loLIM;
   TraceOut_channels_2_bipolar[10] := Binding_7_channels[2].bipolar;
   TraceOut_channels_2_measuringMode[10] := Binding_7_channels[2].measuringMode;
   TraceOut_channels_2_retVal[10] := Binding_7_channels[2].retVal;
   TraceOut_channels_2_outputValue[10] := Binding_7_channels[2].outputValue;
   TraceOut_channels_3_enable[10] := Binding_7_channels[3].enable;
   TraceOut_channels_3_hiLIM[10] := Binding_7_channels[3].hiLIM;
   TraceOut_channels_3_loLIM[10] := Binding_7_channels[3].loLIM;
   TraceOut_channels_3_bipolar[10] := Binding_7_channels[3].bipolar;
   TraceOut_channels_3_measuringMode[10] := Binding_7_channels[3].measuringMode;
   TraceOut_channels_3_retVal[10] := Binding_7_channels[3].retVal;
   TraceOut_channels_3_outputValue[10] := Binding_7_channels[3].outputValue;
   TraceOut_channels_4_enable[10] := Binding_7_channels[4].enable;
   TraceOut_channels_4_hiLIM[10] := Binding_7_channels[4].hiLIM;
   TraceOut_channels_4_loLIM[10] := Binding_7_channels[4].loLIM;
   TraceOut_channels_4_bipolar[10] := Binding_7_channels[4].bipolar;
   TraceOut_channels_4_measuringMode[10] := Binding_7_channels[4].measuringMode;
   TraceOut_channels_4_retVal[10] := Binding_7_channels[4].retVal;
   TraceOut_channels_4_outputValue[10] := Binding_7_channels[4].outputValue;
   TraceOut_channels_5_enable[10] := Binding_7_channels[5].enable;
   TraceOut_channels_5_hiLIM[10] := Binding_7_channels[5].hiLIM;
   TraceOut_channels_5_loLIM[10] := Binding_7_channels[5].loLIM;
   TraceOut_channels_5_bipolar[10] := Binding_7_channels[5].bipolar;
   TraceOut_channels_5_measuringMode[10] := Binding_7_channels[5].measuringMode;
   TraceOut_channels_5_retVal[10] := Binding_7_channels[5].retVal;
   TraceOut_channels_5_outputValue[10] := Binding_7_channels[5].outputValue;
   BenchCalls := BenchCalls + 1;
 11:
   Binding_8_analogValues[1] := INT#-27648;
   Binding_8_analogValues[2] := INT#30000;
   Binding_8_analogValues[3] := INT#-13824;
   Binding_8_analogValues[4] := INT#-255;
   Binding_8_analogValues[5] := INT#12345;
   Binding_8_channels[1].enable := TRUE;
   Binding_8_channels[1].hiLIM := REAL#10.0;
   Binding_8_channels[1].loLIM := REAL#-10.0;
   Binding_8_channels[1].bipolar := TRUE;
   Binding_8_channels[1].measuringMode := INT#0;
   Binding_8_channels[1].retVal := WORD#7;
   Binding_8_channels[1].outputValue := REAL#-999.0;
   Binding_8_channels[2].enable := TRUE;
   Binding_8_channels[2].hiLIM := REAL#100.0;
   Binding_8_channels[2].loLIM := REAL#0.0;
   Binding_8_channels[2].bipolar := FALSE;
   Binding_8_channels[2].measuringMode := INT#0;
   Binding_8_channels[2].retVal := WORD#7;
   Binding_8_channels[2].outputValue := REAL#-999.0;
   Binding_8_channels[3].enable := TRUE;
   Binding_8_channels[3].hiLIM := REAL#100.0;
   Binding_8_channels[3].loLIM := REAL#0.0;
   Binding_8_channels[3].bipolar := FALSE;
   Binding_8_channels[3].measuringMode := INT#0;
   Binding_8_channels[3].retVal := WORD#7;
   Binding_8_channels[3].outputValue := REAL#-999.0;
   Binding_8_channels[4].enable := TRUE;
   Binding_8_channels[4].hiLIM := REAL#100.0;
   Binding_8_channels[4].loLIM := REAL#-100.0;
   Binding_8_channels[4].bipolar := FALSE;
   Binding_8_channels[4].measuringMode := INT#1;
   Binding_8_channels[4].retVal := WORD#7;
   Binding_8_channels[4].outputValue := REAL#-999.0;
   Binding_8_channels[5].enable := TRUE;
   Binding_8_channels[5].hiLIM := REAL#200.0;
   Binding_8_channels[5].loLIM := REAL#-200.0;
   Binding_8_channels[5].bipolar := TRUE;
   Binding_8_channels[5].measuringMode := INT#2;
   Binding_8_channels[5].retVal := WORD#7;
   Binding_8_channels[5].outputValue := REAL#-999.0;
   Binding_8_channels[6].enable := TRUE;
   Binding_8_channels[6].hiLIM := REAL#100.0;
   Binding_8_channels[6].loLIM := REAL#0.0;
   Binding_8_channels[6].bipolar := FALSE;
   Binding_8_channels[6].measuringMode := INT#0;
   Binding_8_channels[6].retVal := WORD#42;
   Binding_8_channels[6].outputValue := REAL#-123.0;
   BenchUut8.count := DINT#5;
   TraceIn_count[11] := BenchUut8.count;
   BenchUut8(analogValues := Binding_8_analogValues, channels := Binding_8_channels);
   TraceOut_analogValues_1[11] := Binding_8_analogValues[1];
   TraceOut_analogValues_2[11] := Binding_8_analogValues[2];
   TraceOut_analogValues_3[11] := Binding_8_analogValues[3];
   TraceOut_analogValues_4[11] := Binding_8_analogValues[4];
   TraceOut_analogValues_5[11] := Binding_8_analogValues[5];
   TraceOut_channels_1_enable[11] := Binding_8_channels[1].enable;
   TraceOut_channels_1_hiLIM[11] := Binding_8_channels[1].hiLIM;
   TraceOut_channels_1_loLIM[11] := Binding_8_channels[1].loLIM;
   TraceOut_channels_1_bipolar[11] := Binding_8_channels[1].bipolar;
   TraceOut_channels_1_measuringMode[11] := Binding_8_channels[1].measuringMode;
   TraceOut_channels_1_retVal[11] := Binding_8_channels[1].retVal;
   TraceOut_channels_1_outputValue[11] := Binding_8_channels[1].outputValue;
   TraceOut_channels_2_enable[11] := Binding_8_channels[2].enable;
   TraceOut_channels_2_hiLIM[11] := Binding_8_channels[2].hiLIM;
   TraceOut_channels_2_loLIM[11] := Binding_8_channels[2].loLIM;
   TraceOut_channels_2_bipolar[11] := Binding_8_channels[2].bipolar;
   TraceOut_channels_2_measuringMode[11] := Binding_8_channels[2].measuringMode;
   TraceOut_channels_2_retVal[11] := Binding_8_channels[2].retVal;
   TraceOut_channels_2_outputValue[11] := Binding_8_channels[2].outputValue;
   TraceOut_channels_3_enable[11] := Binding_8_channels[3].enable;
   TraceOut_channels_3_hiLIM[11] := Binding_8_channels[3].hiLIM;
   TraceOut_channels_3_loLIM[11] := Binding_8_channels[3].loLIM;
   TraceOut_channels_3_bipolar[11] := Binding_8_channels[3].bipolar;
   TraceOut_channels_3_measuringMode[11] := Binding_8_channels[3].measuringMode;
   TraceOut_channels_3_retVal[11] := Binding_8_channels[3].retVal;
   TraceOut_channels_3_outputValue[11] := Binding_8_channels[3].outputValue;
   TraceOut_channels_4_enable[11] := Binding_8_channels[4].enable;
   TraceOut_channels_4_hiLIM[11] := Binding_8_channels[4].hiLIM;
   TraceOut_channels_4_loLIM[11] := Binding_8_channels[4].loLIM;
   TraceOut_channels_4_bipolar[11] := Binding_8_channels[4].bipolar;
   TraceOut_channels_4_measuringMode[11] := Binding_8_channels[4].measuringMode;
   TraceOut_channels_4_retVal[11] := Binding_8_channels[4].retVal;
   TraceOut_channels_4_outputValue[11] := Binding_8_channels[4].outputValue;
   TraceOut_channels_5_enable[11] := Binding_8_channels[5].enable;
   TraceOut_channels_5_hiLIM[11] := Binding_8_channels[5].hiLIM;
   TraceOut_channels_5_loLIM[11] := Binding_8_channels[5].loLIM;
   TraceOut_channels_5_bipolar[11] := Binding_8_channels[5].bipolar;
   TraceOut_channels_5_measuringMode[11] := Binding_8_channels[5].measuringMode;
   TraceOut_channels_5_retVal[11] := Binding_8_channels[5].retVal;
   TraceOut_channels_5_outputValue[11] := Binding_8_channels[5].outputValue;
   TraceOut_channels_6_enable[11] := Binding_8_channels[6].enable;
   TraceOut_channels_6_hiLIM[11] := Binding_8_channels[6].hiLIM;
   TraceOut_channels_6_loLIM[11] := Binding_8_channels[6].loLIM;
   TraceOut_channels_6_bipolar[11] := Binding_8_channels[6].bipolar;
   TraceOut_channels_6_measuringMode[11] := Binding_8_channels[6].measuringMode;
   TraceOut_channels_6_retVal[11] := Binding_8_channels[6].retVal;
   TraceOut_channels_6_outputValue[11] := Binding_8_channels[6].outputValue;
   BenchCalls := BenchCalls + 1;
 END_CASE;
 BenchStep := BenchStep + 1;
 IF BenchStep >= 12 THEN BenchDone := TRUE; END_IF;
END_IF;
END_PROGRAM
